Staubli VAL3: utBorder.pjx

--- utBorder.pjx ---
Parameters version=s8.10Cs9_BS1925 stackSize=5000 millimeterUnit=true
Program file=start.pgx
Program file=stop.pgx
Data file=utBorder.dtx

--- utBorder.dtx ---
public string sBorderColour
public string sBorderSytle
public string sBorderWidth

--- start.pgx ---
program start()
begin
end

--- stop.pgx ---
program stop()
begin
end
